TYPE ST_SetConfigParamParam :
STRUCT
	Id : UDINT;
	DataType : E_ConfigDataType;
	Value : STRING(80);
END_STRUCT
END_TYPE

(* stored: Version 1.1.0.1, ProductVersion 3.1.4026.18
   DUT ST_SetConfigParamParam: Id {8e7b0129-e77b-4814-855f-93745f7990ad} *)
